Staubli VAL3: pointEditValue.pgx

public program pointEditValue(string x_sMoveType, string x_sKey, num x_nIndex, num& x_nTRSF[], string& x_sTRSF[], bool& x_bShow2Point)
begin
  switch x_sMoveType
    case "CIRCLE"
      trajTemp:tTrajItem[x_sKey].pPointItem[x_nIndex].pParaItem.nMoveType=2
      x_nTRSF[0]=trajTemp:tTrajItem[x_sKey].pPointItem[x_nIndex].pPointRx.trsf.x
      x_nTRSF[1]=trajTemp:tTrajItem[x_sKey].pPointItem[x_nIndex].pPointRx.trsf.y
      x_nTRSF[2]=trajTemp:tTrajItem[x_sKey].pPointItem[x_nIndex].pPointRx.trsf.z
      x_nTRSF[3]=trajTemp:tTrajItem[x_sKey].pPointItem[x_nIndex].pPointRx.trsf.rx
      x_nTRSF[4]=trajTemp:tTrajItem[x_sKey].pPointItem[x_nIndex].pPointRx.trsf.ry
      x_nTRSF[5]=trajTemp:tTrajItem[x_sKey].pPointItem[x_nIndex].pPointRx.trsf.rz
      x_nTRSF[6]=trajTemp:tTrajItem[x_sKey].pPointItem[x_nIndex].pInter.trsf.x
      x_nTRSF[7]=trajTemp:tTrajItem[x_sKey].pPointItem[x_nIndex].pInter.trsf.y
      x_nTRSF[8]=trajTemp:tTrajItem[x_sKey].pPointItem[x_nIndex].pInter.trsf.z
      x_nTRSF[9]=trajTemp:tTrajItem[x_sKey].pPointItem[x_nIndex].pInter.trsf.rx
      x_nTRSF[10]=trajTemp:tTrajItem[x_sKey].pPointItem[x_nIndex].pInter.trsf.ry
      x_nTRSF[11]=trajTemp:tTrajItem[x_sKey].pPointItem[x_nIndex].pInter.trsf.rz
      x_sTRSF[0]="X:"
      x_sTRSF[1]="Y:"
      x_sTRSF[2]="Z:"
      x_sTRSF[3]="RX:"
      x_sTRSF[4]="RY:"
      x_sTRSF[5]="RZ:"
      x_sTRSF[6]="2X:"
      x_sTRSF[7]="2Y:"
      x_sTRSF[8]="2Z:"
      x_sTRSF[9]="2RX:"
      x_sTRSF[10]="2RY:"
      x_sTRSF[11]="2RZ:"
      x_bShow2Point=true
    break
    case "POINT"
      trajTemp:tTrajItem[x_sKey].pPointItem[x_nIndex].pParaItem.nMoveType=1
      x_nTRSF[0]=trajTemp:tTrajItem[x_sKey].pPointItem[x_nIndex].pPointRx.trsf.x
      x_nTRSF[1]=trajTemp:tTrajItem[x_sKey].pPointItem[x_nIndex].pPointRx.trsf.y
      x_nTRSF[2]=trajTemp:tTrajItem[x_sKey].pPointItem[x_nIndex].pPointRx.trsf.z
      x_nTRSF[3]=trajTemp:tTrajItem[x_sKey].pPointItem[x_nIndex].pPointRx.trsf.rx
      x_nTRSF[4]=trajTemp:tTrajItem[x_sKey].pPointItem[x_nIndex].pPointRx.trsf.ry
      x_nTRSF[5]=trajTemp:tTrajItem[x_sKey].pPointItem[x_nIndex].pPointRx.trsf.rz
      x_sTRSF[0]="X:"
      x_sTRSF[1]="Y:"
      x_sTRSF[2]="Z:"
      x_sTRSF[3]="RX:"
      x_sTRSF[4]="RY:"
      x_sTRSF[5]="RZ:"
    break
    case "JOINT"
      trajTemp:tTrajItem[x_sKey].pPointItem[x_nIndex].pParaItem.nMoveType=0
      x_nTRSF[0]=trajTemp:tTrajItem[x_sKey].pPointItem[x_nIndex].jJointRx.j1
      x_nTRSF[1]=trajTemp:tTrajItem[x_sKey].pPointItem[x_nIndex].jJointRx.j2
      x_nTRSF[2]=trajTemp:tTrajItem[x_sKey].pPointItem[x_nIndex].jJointRx.j3
      x_nTRSF[3]=trajTemp:tTrajItem[x_sKey].pPointItem[x_nIndex].jJointRx.j4
      x_nTRSF[4]=trajTemp:tTrajItem[x_sKey].pPointItem[x_nIndex].jJointRx.j5
      x_nTRSF[5]=trajTemp:tTrajItem[x_sKey].pPointItem[x_nIndex].jJointRx.j6
      x_sTRSF[0]="J1:"
      x_sTRSF[1]="J2:"
      x_sTRSF[2]="J3:"
      x_sTRSF[3]="J4:"
      x_sTRSF[4]="J5:"
      x_sTRSF[5]="J6:"
    break
  endSwitch
end
